SUBAPPLICATION Uebung_260_AX (* Frequenzgenerator: Poti I1 0..100 % = 0..1000 Hz (mHz) auf Q1, Tastgrad 50 % *)
  (* Standard: 61499-2; Description: Copyright (c) 2026 Meisterschulen am Ostbahnhof This program and the accompanying materials are made available under the terms of the Eclipse Public License 2.0 which is available at https://www.eclipse.org/legal/epl-2.0/ SPDX-License-Identifier: EPL-2.0 *)
  (* Version 1.0, 2026-11-06, Franz Höpfinger, Meisterschulen am Ostbahnhof, initial API and implementation and/or initial documentation *)
  PACKAGE Uebungen;
  IMPORT logiBUS::io::AI::logiBUS_AI::AnalogInput_I1;
  IMPORT Meins::InputOutputTester::Button_AI_Calibrate_2P_OPC_UA::SubStrings::AIC_I1_RAW_WRITE;
  IMPORT Meins::InputOutputTester::Button_AI_Calibrate_2P_OPC_UA::SubStrings::AIC_I1_CAL_WRITE;
  IMPORT Meins::InputOutputTester::Button_AI_Calibrate_2P_OPC_UA::SubStrings::AIC_I1_CO_METHOD;
  IMPORT Meins::InputOutputTester::Button_AI_Calibrate_2P_OPC_UA::SubStrings::AIC_I1_CS_METHOD;
  IMPORT Meins::InputOutputTester::Button_AI_Calibrate_2P_OPC_UA::SubStrings::AIC_I1_ZERO_READ;
  IMPORT Meins::InputOutputTester::Button_AI_Calibrate_2P_OPC_UA::SubStrings::AIC_I1_ZERO_WRITE;
  IMPORT Meins::InputOutputTester::Button_AI_Calibrate_2P_OPC_UA::SubStrings::AIC_I1_SPAN_READ;
  IMPORT Meins::InputOutputTester::Button_AI_Calibrate_2P_OPC_UA::SubStrings::AIC_I1_SPAN_WRITE;
  IMPORT Meins::InputOutputTester::Button_AI_Calibrate_2P_OPC_UA::SubStrings::AIC_I1_ZERO_RAW_WRITE;
  IMPORT Meins::InputOutputTester::Button_AI_Calibrate_2P_OPC_UA::SubStrings::AIC_I1_SPAN_RAW_WRITE;
  IMPORT logiBUS::io::DQ::logiBUS_DO::Output_Q1;
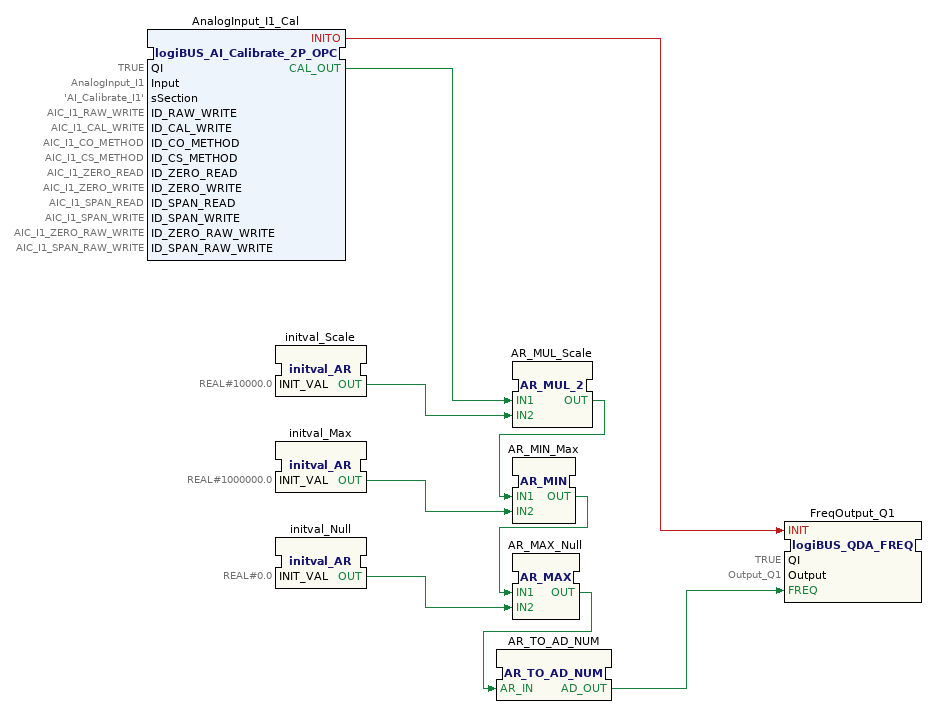
  (* Vorher AI1 kalibrieren: 1. Meins/InputOutputTester/Button_AI_Calibrate_2P_OPC_UA als Control in test_AX.sys, Bootfile exportieren, aufspielen. 2. Mit Web-Clients/apixon-ai-calibrate-2p-client/dist/apixon-ai-calibrate-2p.html AI1 kalibrieren (0 %: CO, 100 %: CS). 3. INI-Datei auf der Platine liegen lassen (Sektion AI_Calibrate_I1). Danach laeuft diese Uebung ohne VT und ohne Dashboard. *)
  FBS
    AR_MUL_Scale : adapter::iec61131::arithmetic::AR_MUL_2;
    initval_Scale : adapter::types::unidirectional::AR::initval::initval_AR(INIT_VAL := REAL#10000.0);
    AR_MIN_Max : adapter::iec61131::selection::AR_MIN;
    initval_Max : adapter::types::unidirectional::AR::initval::initval_AR(INIT_VAL := REAL#1000000.0);
    AR_MAX_Null : adapter::iec61131::selection::AR_MAX;
    initval_Null : adapter::types::unidirectional::AR::initval::initval_AR(INIT_VAL := REAL#0.0);
    AR_TO_AD_NUM : adapter::conversion::unidirectional::AR_TO_AD_NUM;
    FreqOutput_Q1 : logiBUS::io::DQ::logiBUS_QDA_FREQ(QI := TRUE, Output := Output_Q1);
  END_FBS
  SUBAPPS
    AnalogInput_I1_Cal : MyLib::sys::logiBUS_AI_Calibrate_2P_OPC(QI := TRUE, Input := AnalogInput_I1, sSection := 'AI_Calibrate_I1', ID_RAW_WRITE := AIC_I1_RAW_WRITE, ID_CAL_WRITE := AIC_I1_CAL_WRITE, ID_CO_METHOD := AIC_I1_CO_METHOD, ID_CS_METHOD := AIC_I1_CS_METHOD, ID_ZERO_READ := AIC_I1_ZERO_READ, ID_ZERO_WRITE := AIC_I1_ZERO_WRITE, ID_SPAN_READ := AIC_I1_SPAN_READ, ID_SPAN_WRITE := AIC_I1_SPAN_WRITE, ID_ZERO_RAW_WRITE := AIC_I1_ZERO_RAW_WRITE, ID_SPAN_RAW_WRITE := AIC_I1_SPAN_RAW_WRITE);
  END_SUBAPPS
  EVENT_CONNECTIONS
    AnalogInput_I1_Cal.INITO TO FreqOutput_Q1.INIT;
  END_CONNECTIONS
  ADAPTER_CONNECTIONS
    AnalogInput_I1_Cal.CAL_OUT TO AR_MUL_Scale.IN1;
    initval_Scale.OUT TO AR_MUL_Scale.IN2;
    AR_MUL_Scale.OUT TO AR_MIN_Max.IN1;
    initval_Max.OUT TO AR_MIN_Max.IN2;
    AR_MIN_Max.OUT TO AR_MAX_Null.IN1;
    initval_Null.OUT TO AR_MAX_Null.IN2;
    AR_MAX_Null.OUT TO AR_TO_AD_NUM.AR_IN;
    AR_TO_AD_NUM.AD_OUT TO FreqOutput_Q1.FREQ;
  END_CONNECTIONS
END_SUBAPPLICATION
